Fanuc KAREL source: kb00039.KL

-- PROVISIONAL review KL for V940-1; original PC SHA256 1664f8c3b2274f7528a082960226b047fe6566fb6121422c5cc0a4eb2f39763b
-- Incomplete behavior may be omitted. Consult companion uncertainty JSON. Do not deploy.
PROGRAM KB00039
%NOLOCKGROUP
BEGIN
  -- V9_ZERO_TABLE_METADATA_HINT layout=0002_ascii; no indexed target words; source/name/runtime held
  -- UNRESOLVED_PC offsets 5-14; opcodes 3F,75
  -- UNRESOLVED_PC offsets 19-26; opcodes 9D,23
  -- UNRESOLVED_PC offsets 31-55; opcodes 27,22,2A,22,22,31
  -- UNRESOLVED_PC offsets 60-64; opcodes 7F
END KB00039
